Fanuc KAREL source: KT00630.KL

PROGRAM KT00630
%NOLOCKGROUP
VAR
  S1: STRING[80]
  S2: STRING[80]
  OUT: BOOLEAN
BEGIN
  S1 = 'A'
  S2 = 'B'
  S1 = 'A'
  S2 = 'B'
  OUT = + S1
END KT00630
